Fanuc KAREL source: kb00053.KL

PROGRAM KB00053
%STACKSIZE=65535
%PRIORITY=65535
%NOLOCKGROUP
VAR
RESULT : STRING[80]
BEGIN
RESULT=CURR_PROG()
END KB00053
